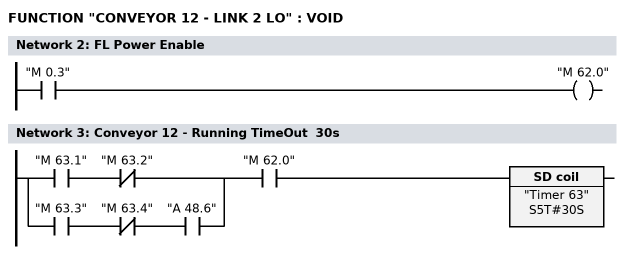

      A     "M 0.3";
      =     "M 62.0";
NETWORK
TITLE =Conveyor 12 - Running TimeOut  30s

      A(    ;
      A     "M 63.1";
      AN    "M 63.2";
      O     ;
      A     "M 63.3";
      AN    "M 63.4";
      A     "A 48.6";
      )     ;
      A     "M 62.0";
      L     S5T#30S;
      SD    "Timer 63";
NETWORK
TITLE =Conveyor 12 - Steps Register - Reset

      A(    ;
      A     "M 63.1";
      AN    "M 63.2";
      A     "Timer 63";
      O     "M 63.4";
      )     ;
      A     "M 62.0";
      JC    M001;
      JU    M002;

M001: L     W#16#0;
      T     "MW 63";
      T     "MB 65";

M002: NOP   0;
NETWORK
TITLE =Step 13N1 - Power On
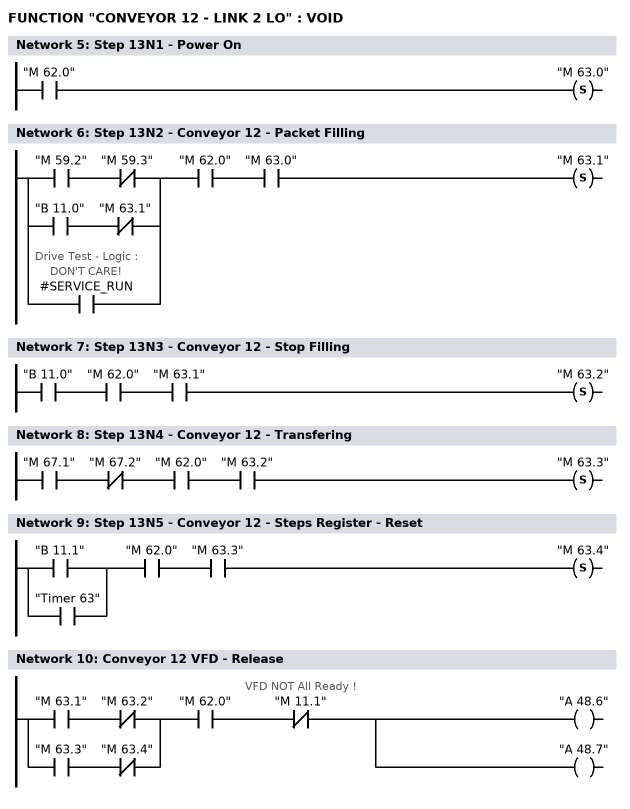

      A     "M 62.0";
      S     "M 63.0";
NETWORK
TITLE =Step 13N2 - Conveyor 12 - Packet Filling

      A(    ;
      A     "M 59.2";
      AN    "M 59.3";
      O     ;
      A     "B 11.0";
      AN    "M 63.1";
      )     ;
      O     #SERVICE_RUN; // Drive Test - Logic : DON'T CARE!
      A     "M 62.0";
      A     "M 63.0";
      S     "M 63.1";
NETWORK
TITLE =Step 13N3 - Conveyor 12 - Stop Filling

      A     "B 11.0";
      A     "M 62.0";
      A     "M 63.1";
      S     "M 63.2";
NETWORK
TITLE =Step 13N4 - Conveyor 12 - Transfering

      A     "M 67.1";
      AN    "M 67.2";
      A     "M 62.0";
      A     "M 63.2";
      S     "M 63.3";
NETWORK
TITLE =Step 13N5 - Conveyor 12 - Steps Register - Reset

      A(    ;
      O     "B 11.1";
      O     "Timer 63";
      )     ;
      A     "M 62.0";
      A     "M 63.3";
      S     "M 63.4";
NETWORK
TITLE =Conveyor 12 VFD - Release

      A(    ;
      A     "M 63.1";
      AN    "M 63.2";
      O     ;
      A     "M 63.3";
      AN    "M 63.4";
      )     ;
      A     "M 62.0";
      AN    "M 11.1"; // VFD NOT All Ready !
      =     "A 48.6";
      =     "A 48.7";
END_FUNCTION

FUNCTION "CONVEYOR 13 - DELIV. LO" : VOID
TITLE =Conveyor 13 - Delivery First Level
NAME : POS_15_L
VERSION : 0.0


VAR_TEMP
  MAIN_SERVICE_2_SW : BOOL ;
  SERVICE_RUN : BOOL ;
  BARRIER_BLINKER : BOOL ;	//Feeder Safety Light Barrier
END_VAR
BEGIN
NETWORK
TITLE =Conveyor 13 - Service

      A     "HMI_DB".ALL_SERVICE_ENABLE_SW;
      A     "HMI_DB".CONVEYOR_11_SERVICE_SW;
      A     "HMI_DB".SERVICE_SW_2_STATUS;
      =     #MAIN_SERVICE_2_SW;
//;
      A     #MAIN_SERVICE_2_SW;
      O     "M 66.1";
      JNB   CO13;
//;
      A     "HMI_DB".HMI_CONVEYOR_13_TEST_SSW;
      =     #SERVICE_RUN;
//;
      AN    #MAIN_SERVICE_2_SW;
      R     "HMI_DB".HMI_CONVEYOR_13_TEST_SSW;

CO13: R     #SERVICE_RUN;
      FP    "FP 148.2";
      =     "M 66.1";
NETWORK
TITLE =Delivery Conveyor 13 - Running TimeOut  30s
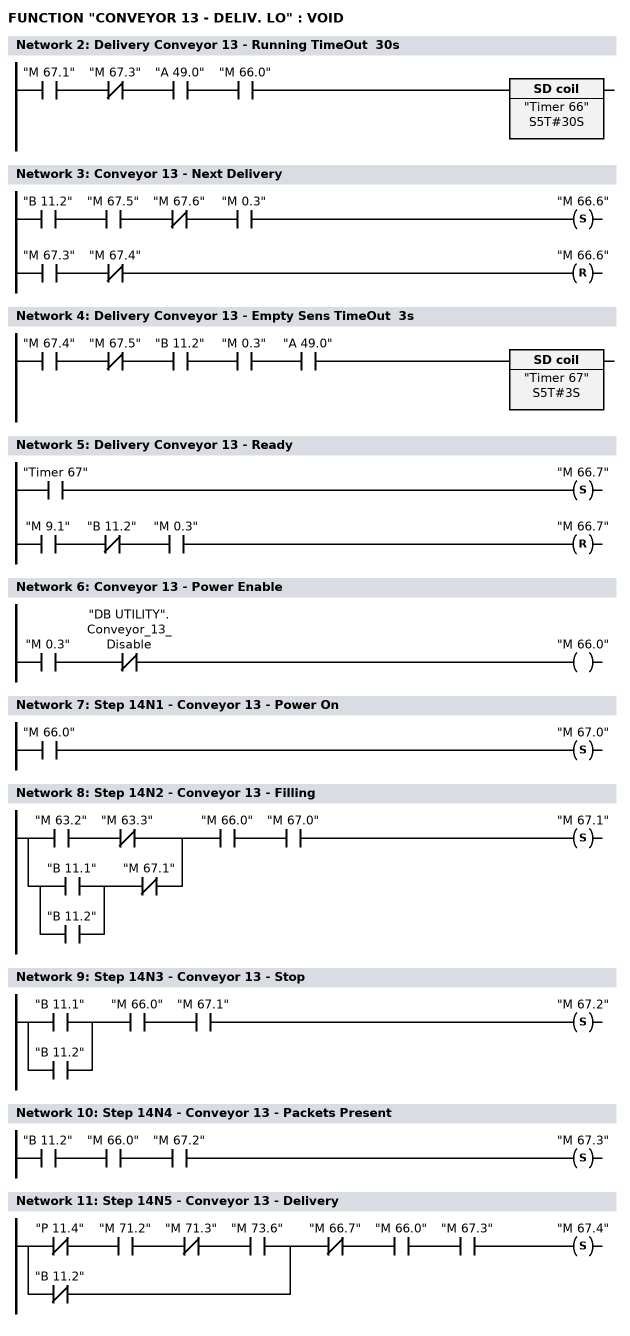

      A     "M 67.1";
      AN    "M 67.3";
      A     "A 49.0";
      A     "M 66.0";
      L     S5T#30S;
      SD    "Timer 66";
NETWORK
TITLE =Conveyor 13 - Next Delivery

      A     "B 11.2";
      A     "M 67.5";
      AN    "M 67.6";
      A     "M 0.3";
      S     "M 66.6";
//;
      A     "M 67.3";
      AN    "M 67.4";
      R     "M 66.6";
NETWORK
TITLE =Delivery Conveyor 13 - Empty Sens TimeOut  3s

      A     "M 67.4";
      AN    "M 67.5";
      A     "B 11.2";
      A     "M 0.3";
      A     "A 49.0";
      L     S5T#3S;
      SD    "Timer 67";
NETWORK
TITLE =Delivery Conveyor 13 - Ready

      A     "Timer 67";
      S     "M 66.7";
//;
      A     "M 9.1";
      AN    "B 11.2";
      A     "M 0.3";
      R     "M 66.7";
NETWORK
TITLE =Conveyor 13 - Power Enable

      A     "M 0.3";
      AN    "DB UTILITY".Conveyor_13_Disable;
      =     "M 66.0";
NETWORK
TITLE =Step 14N1 - Conveyor 13 - Power On

      A     "M 66.0";
      S     "M 67.0";
NETWORK
TITLE =Step 14N2 - Conveyor 13 - Filling

      A(    ;
      A     "M 63.2";
      AN    "M 63.3";
      O     ;
      A(    ;
      O     "B 11.1";
      O     "B 11.2";
      )     ;
//      O     #SERVICE_RUN
      AN    "M 67.1";
      )     ;
      A     "M 66.0";
      A     "M 67.0";
      S     "M 67.1";
NETWORK
TITLE =Step 14N3 - Conveyor 13 - Stop

      A(    ;
      O     "B 11.1";
      O     "B 11.2";
      )     ;
      A     "M 66.0";
      A     "M 67.1";
      S     "M 67.2";
NETWORK
TITLE =Step 14N4 - Conveyor 13 - Packets Present

      A     "B 11.2";
      A     "M 66.0";
      A     "M 67.2";
      S     "M 67.3";
NETWORK
TITLE =Step 14N5 - Conveyor 13 - Delivery

      A(    ;
      AN    "P 11.4";
      A     "M 71.2";
      AN    "M 71.3";
      A     "M 73.6";
      ON    "B 11.2";
      )     ;
      AN    "M 66.7";
      A     "M 66.0";
      A     "M 67.3";
      S     "M 67.4";
NETWORK
TITLE =Write 1 to Steps 0-3 Byte Register MB67

      A(    ;
      O     "M 66.6";
      O     "M 66.7";
      )     ;
      A     "M 67.4";
      A     "M 66.0";
      JC    M001;
      JU    M002;

M001: L     2#1111;
      T     "MB 67";

M002: NOP   0;
NETWORK
TITLE =Step 14N6 - Conveyor 13 - Delivery Done
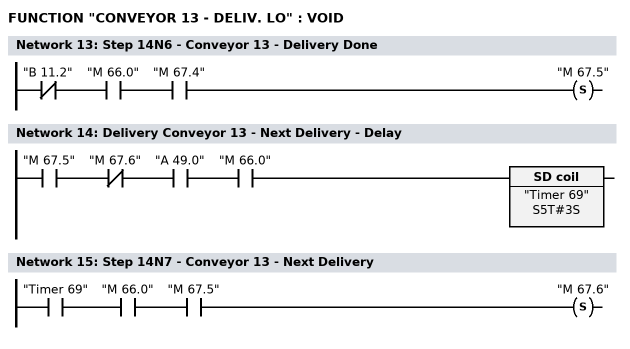

      AN    "B 11.2";
      A     "M 66.0";
      A     "M 67.4";
      S     "M 67.5";
NETWORK
TITLE =Delivery Conveyor 13 - Next Delivery - Delay

      A     "M 67.5";
      AN    "M 67.6";
      A     "A 49.0";
      A     "M 66.0";
      L     S5T#3S;
      SD    "Timer 69";
NETWORK
TITLE =Step 14N7 - Conveyor 13 - Next Delivery

      A     "Timer 69";
      A     "M 66.0";
      A     "M 67.5";
      S     "M 67.6";
NETWORK
TITLE =Steps Register - Reset

      A(    ;
      O     "M 67.6";
      O     "Timer 66";
      )     ;
      A     "M 66.0";
      JC    M003;
      JU    M004;

M003: L     2#0;
      T     "MW 67";

M004: NOP   0;
NETWORK
TITLE =Conveyor 13 VFD - Release
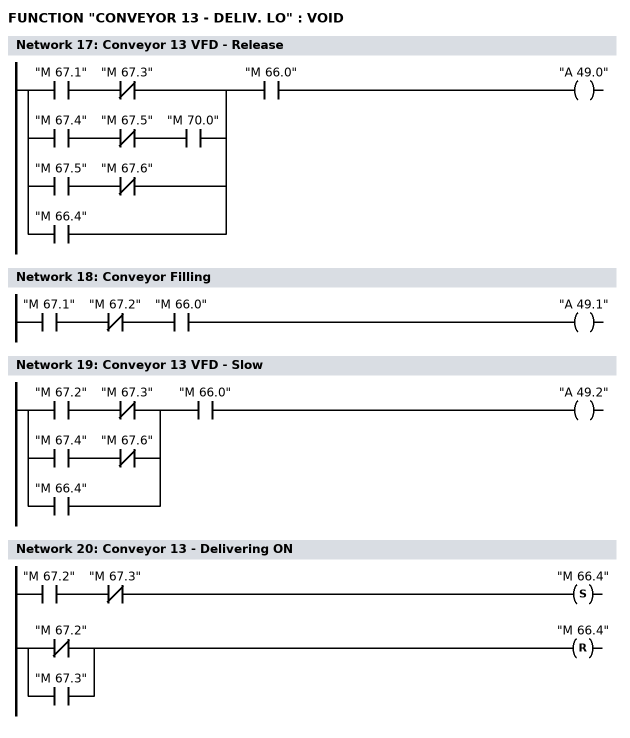

      A(    ;
      A     "M 67.1";
      AN    "M 67.3";
      O     ;
      A     "M 67.4";
      AN    "M 67.5";
      A     "M 70.0";
      O     ;
      A     "M 67.5";
      AN    "M 67.6";
      O     "M 66.4";
      )     ;
      A     "M 66.0";
      =     "A 49.0";
NETWORK
TITLE =Conveyor Filling

      A     "M 67.1";
      AN    "M 67.2";
      A     "M 66.0";
      =     "A 49.1";
NETWORK
TITLE =Conveyor 13 VFD - Slow

      A(    ;
      A     "M 67.2";
      AN    "M 67.3";
      O     ;
      A     "M 67.4";
      AN    "M 67.6";
      O     "M 66.4";
      )     ;
      A     "M 66.0";
      =     "A 49.2";
NETWORK
TITLE =Conveyor 13 - Delivering ON

      A     "M 67.2";
      AN    "M 67.3";
      S     "M 66.4";
//;
      A(    ;
      ON    "M 67.2";
      O     "M 67.3";
      )     ;
      R     "M 66.4";
END_FUNCTION

FUNCTION "LOADER FINGERS" : VOID
TITLE =Feeder Fingers
//
NAME : FEEDER
VERSION : 0.0


VAR_TEMP
  MAIN_SERVICE_3_SW : BOOL ;
  FEEDER_SERVICE_SW : BOOL ;
  FINGERS_SERVICE_SW : BOOL ;
  LIGHT_BARRIER : BOOL ;
  FINGERS_EXTEND : BOOL ;
  FINGERS_RETRACT : BOOL ;
  FINGERS_TILT : BOOL ;
  BELT_ON : BOOL ;
  INITIALISATION : BOOL ;
END_VAR
BEGIN
NETWORK
TITLE =Light Barrier Buffer
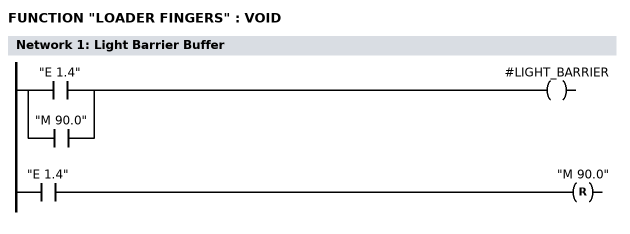

      A     "E 1.4";
      O     "M 90.0";
      =     #LIGHT_BARRIER;
//;
      A     "E 1.4";
      R     "M 90.0";
NETWORK
TITLE =Feeder Service

      A     "HMI_DB".ALL_SERVICE_ENABLE_SW;
      A     "HMI_DB".LOADER_SERVICE_ENABLE_SW;
      A     "HMI_DB".SERVICE_SW_3_STATUS;
      =     #MAIN_SERVICE_3_SW;
//;
      A     #MAIN_SERVICE_3_SW;
      O     "M 70.7";
      JNB   FEED;
      A     "HMI_DB".LOADER_LIFT_SERVICE_SSW;
      =     #FEEDER_SERVICE_SW;
//;
      A     #FEEDER_SERVICE_SW;
      A     "HMI_DB".LOADER_FING_SERVICE_SSW;
      =     #FINGERS_SERVICE_SW;
      =     "DB UTILITY".Conveyor_13_Disable;
      =     "DB UTILITY".Conveyor_23_Disable;
//;
      A     #FEEDER_SERVICE_SW;
      A     #FINGERS_SERVICE_SW;
      A     "HMI_DB".FINGER_EXTEND_TEST_PB;
      AN    #FINGERS_RETRACT;
      =     #FINGERS_EXTEND;
//;
      A     #FEEDER_SERVICE_SW;
      A     #FINGERS_SERVICE_SW;
      A     "HMI_DB".FINGER_RETRACT_TEST_PB;
      AN    #FINGERS_EXTEND;
      =     #FINGERS_RETRACT;
//;
      A     #FEEDER_SERVICE_SW;
      A     #FINGERS_SERVICE_SW;
      A     "HMI_DB".FINGER_BELT_TEST_SW;
      =     #BELT_ON;
//;
      A     #FEEDER_SERVICE_SW;
      A     #FINGERS_SERVICE_SW;
      A     "HMI_DB".FINGER_TILT_TEST_PB;
      =     #FINGERS_TILT;
//;
      AN    #MAIN_SERVICE_3_SW;
      ON    #FEEDER_SERVICE_SW;
      R     "HMI_DB".LOADER_FING_SERVICE_SSW;
      R     "HMI_DB".LOADER_LIFT_SERVICE_SSW;
      R     "HMI_DB".FINGER_RETRACT_TEST_PB;
      R     "HMI_DB".FINGER_EXTEND_TEST_PB;
      R     "HMI_DB".FINGER_TILT_TEST_PB;
      R     "HMI_DB".FINGER_BELT_TEST_SW;

FEED: R     #FEEDER_SERVICE_SW;
      R     #FINGERS_SERVICE_SW;
      R     #FINGERS_EXTEND;
      R     #FINGERS_RETRACT;
      R     #FINGERS_TILT;
      FP    "FP 159.7";
      =     "M 70.7";
//;
      A     "HMI_DB".SERVICE_INIT_PB;
      A     #FEEDER_SERVICE_SW;
      A     #MAIN_SERVICE_3_SW;
      =     #INITIALISATION;
NETWORK
TITLE =Feeder - Power Enable
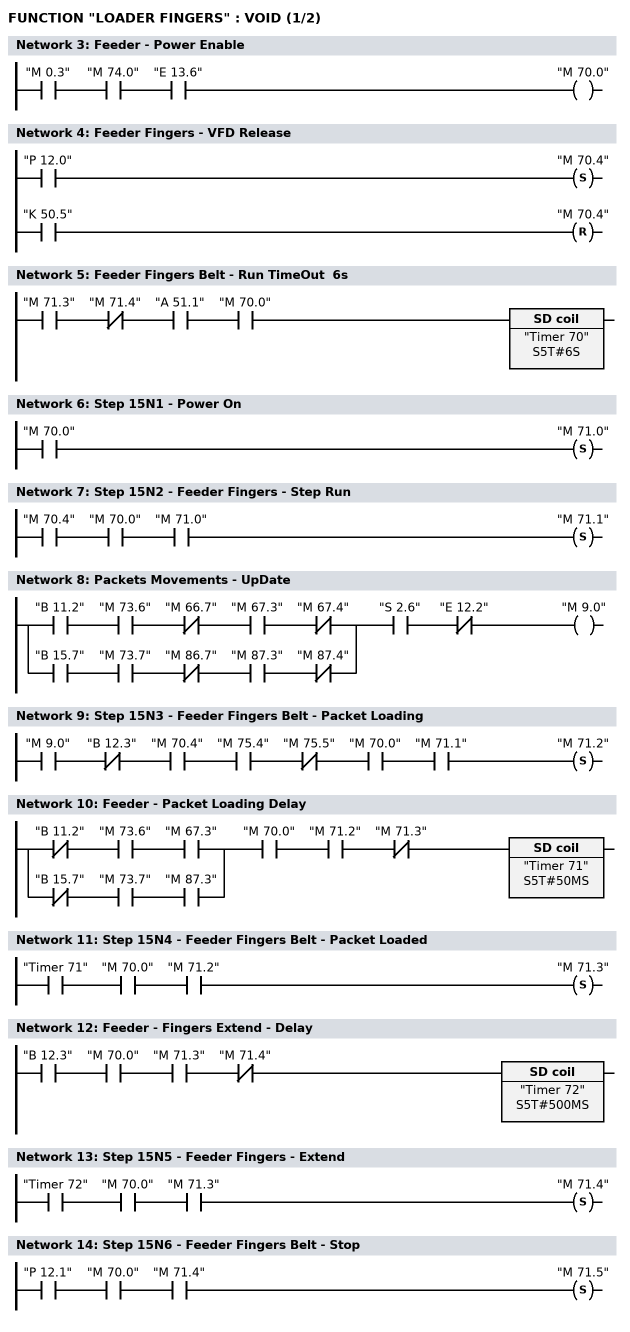

      A     "M 0.3";
      A     "M 74.0";
      A     "E 13.6";
      =     "M 70.0";
NETWORK
TITLE =Feeder Fingers - VFD Release

      A     "P 12.0";
      S     "M 70.4";
//;
      A     "K 50.5";
      R     "M 70.4";
NETWORK
TITLE =Feeder Fingers Belt - Run TimeOut  6s

      A     "M 71.3";
      AN    "M 71.4";
      A     "A 51.1";
      A     "M 70.0";
      L     S5T#6S;
      SD    "Timer 70";
NETWORK
TITLE =Step 15N1 - Power On

      A     "M 70.0";
      S     "M 71.0";
NETWORK
TITLE =Step 15N2 - Feeder Fingers - Step Run

      A     "M 70.4";
      A     "M 70.0";
      A     "M 71.0";
      S     "M 71.1";
NETWORK
TITLE =Packets Movements - UpDate

      A(    ;
      A     "B 11.2";
      A     "M 73.6";
      AN    "M 66.7";
      A     "M 67.3";
      AN    "M 67.4";
      O     ;
      A     "B 15.7";
      A     "M 73.7";
      AN    "M 86.7";
      A     "M 87.3";
      AN    "M 87.4";
      )     ;
      A     "S 2.6";
      AN    "E 12.2";
      =     "M 9.0";
NETWORK
TITLE =Step 15N3 - Feeder Fingers Belt - Packet Loading

      A     "M 9.0";
      AN    "B 12.3";
      A     "M 70.4";
      A     "M 75.4";
      AN    "M 75.5";
      A     "M 70.0";
      A     "M 71.1";
      S     "M 71.2";
NETWORK
TITLE =Feeder - Packet Loading Delay

      A(    ;
      AN    "B 11.2";
      A     "M 73.6";
      A     "M 67.3";
      O     ;
      AN    "B 15.7";
      A     "M 73.7";
      A     "M 87.3";
      )     ;
      A     "M 70.0";
      A     "M 71.2";
      AN    "M 71.3";
      L     S5T#50MS;
      SD    "Timer 71";
NETWORK
TITLE =Step 15N4 - Feeder Fingers Belt - Packet Loaded

      A     "Timer 71";
      A     "M 70.0";
      A     "M 71.2";
      S     "M 71.3";
NETWORK
TITLE =Feeder - Fingers Extend - Delay

      A     "B 12.3";
      A     "M 70.0";
      A     "M 71.3";
      AN    "M 71.4";
      L     S5T#500MS;
      SD    "Timer 72";
NETWORK
TITLE =Step 15N5 - Feeder Fingers - Extend

      A     "Timer 72";
      A     "M 70.0";
      A     "M 71.3";
      S     "M 71.4";
NETWORK
TITLE =Step 15N6 - Feeder Fingers Belt - Stop

      A     "P 12.1";
      A     "M 70.0";
      A     "M 71.4";
      S     "M 71.5";
NETWORK
TITLE =Step 15N7 - Feeder Fingers Tilt - Ready
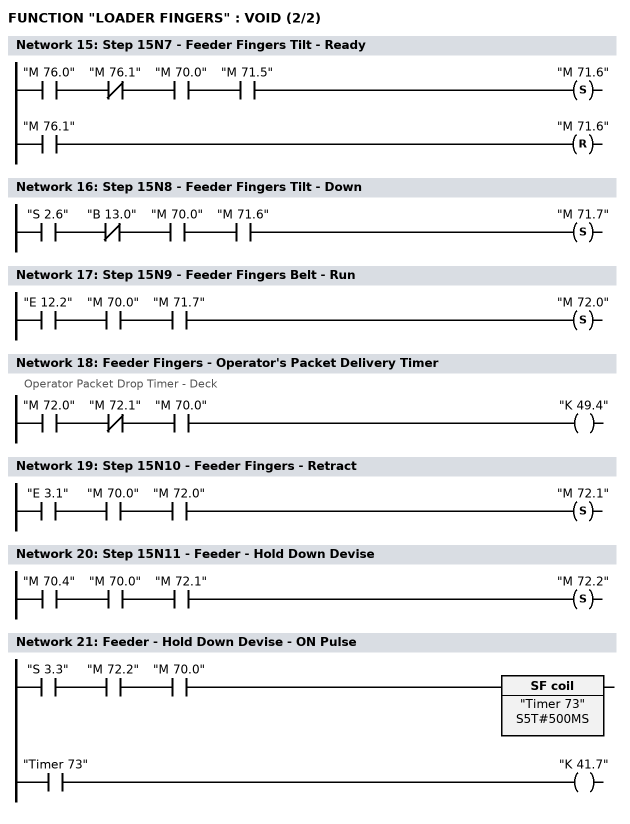

      A     "M 76.0";
      AN    "M 76.1";
      A     "M 70.0";
      A     "M 71.5";
      S     "M 71.6";
//;
      O     "M 76.1";
      R     "M 71.6";
NETWORK
TITLE =Step 15N8 - Feeder Fingers Tilt - Down

      A     "S 2.6";
      AN    "B 13.0";
      A     "M 70.0";
      A     "M 71.6";
      S     "M 71.7";
NETWORK
TITLE =Step 15N9 - Feeder Fingers Belt - Run

      A     "E 12.2";
      A     "M 70.0";
      A     "M 71.7";
      S     "M 72.0";
NETWORK
TITLE =Feeder Fingers - Operator's Packet Delivery Timer
//Operator Packet Drop Timer - Deck
      A     "M 72.0";
      AN    "M 72.1";
      A     "M 70.0";
      =     "K 49.4";
NETWORK
TITLE =Step 15N10 - Feeder Fingers - Retract

      A     "E 3.1";
      A     "M 70.0";
      A     "M 72.0";
      S     "M 72.1";
NETWORK
TITLE =Step 15N11 - Feeder - Hold Down Devise

      A     "M 70.4";
      A     "M 70.0";
      A     "M 72.1";
      S     "M 72.2";
NETWORK
TITLE =Feeder - Hold Down Devise - ON Pulse

      A     "S 3.3";
      A     "M 72.2";
      A     "M 70.0";
      L     S5T#500MS;
      SF    "Timer 73";

      A     "Timer 73";
      =     "K 41.7";
NETWORK
TITLE =Feeder Fingers - Steps Chain Register Reset

      A(    ;
      ON    "M 75.0";
      O     "M 72.2";
      O     "Timer 70";
      O     #FEEDER_SERVICE_SW;
      )     ;
      JC    M001;
      JU    M002;

M001: L     2#0;
      T     "MW 71";

M002: NOP   0;
NETWORK
TITLE =Feeder Fingers - Fingers Retract
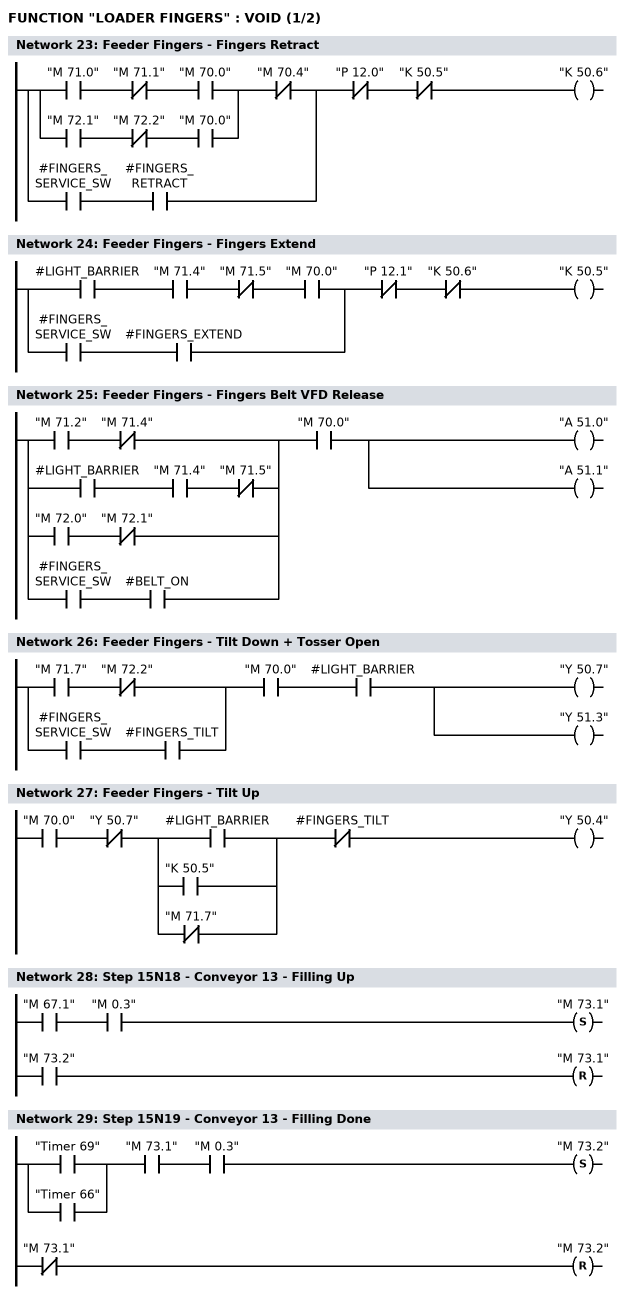

      A(    ;
      A(    ;
      A     "M 71.0";
      AN    "M 71.1";
      A     "M 70.0";
      O     ;
      A     "M 72.1";
      AN    "M 72.2";
      A     "M 70.0";
      )     ;
      AN    "M 70.4";
      O     ;
      A     #FINGERS_SERVICE_SW;
      A     #FINGERS_RETRACT;
      )     ;
      AN    "P 12.0";
      AN    "K 50.5";
      =     "K 50.6";
NETWORK
TITLE =Feeder Fingers - Fingers Extend

      A(    ;
      A     #LIGHT_BARRIER;
      A     "M 71.4";
      AN    "M 71.5";
      A     "M 70.0";
      O     ;
      A     #FINGERS_SERVICE_SW;
      A     #FINGERS_EXTEND;
      )     ;
      AN    "P 12.1";
      AN    "K 50.6";
      =     "K 50.5";
NETWORK
TITLE =Feeder Fingers - Fingers Belt VFD Release

      A(    ;
      A     "M 71.2";
      AN    "M 71.4";
      O     ;
      A     #LIGHT_BARRIER;
      A     "M 71.4";
      AN    "M 71.5";
      O     ;
      A     "M 72.0";
      AN    "M 72.1";
      O     ;
      A     #FINGERS_SERVICE_SW;
      A     #BELT_ON;
      )     ;
      A     "M 70.0";
      =     "A 51.0";
      =     "A 51.1";
NETWORK
TITLE =Feeder Fingers - Tilt Down + Tosser Open

      A(    ;
      A     "M 71.7";
      AN    "M 72.2";
      O     ;
      A     #FINGERS_SERVICE_SW;
      A     #FINGERS_TILT;
      )     ;
      A     "M 70.0";
      A     #LIGHT_BARRIER;
      =     "Y 50.7";
      =     "Y 51.3";
NETWORK
TITLE =Feeder Fingers - Tilt Up

      A     "M 70.0";
      AN    "Y 50.7";
      A(    ;
      O     #LIGHT_BARRIER;
      O     "K 50.5";
      ON    "M 71.7";
      AN    #FINGERS_TILT;
      )     ;
      =     "Y 50.4";
NETWORK
TITLE =Step 15N18 - Conveyor 13 - Filling Up

      A     "M 67.1";
      A     "M 0.3";
      S     "M 73.1";
//;
      A     "M 73.2";
      R     "M 73.1";
NETWORK
TITLE =Step 15N19 - Conveyor 13 - Filling Done

      A(    ;
      O     "Timer 69";
      O     "Timer 66";
      )     ;
      A     "M 73.1";
      A     "M 0.3";
      S     "M 73.2";
//;
      AN    "M 73.1";
      R     "M 73.2";
NETWORK
TITLE =Step 15N20 - Conveyor 23 - Filling Up
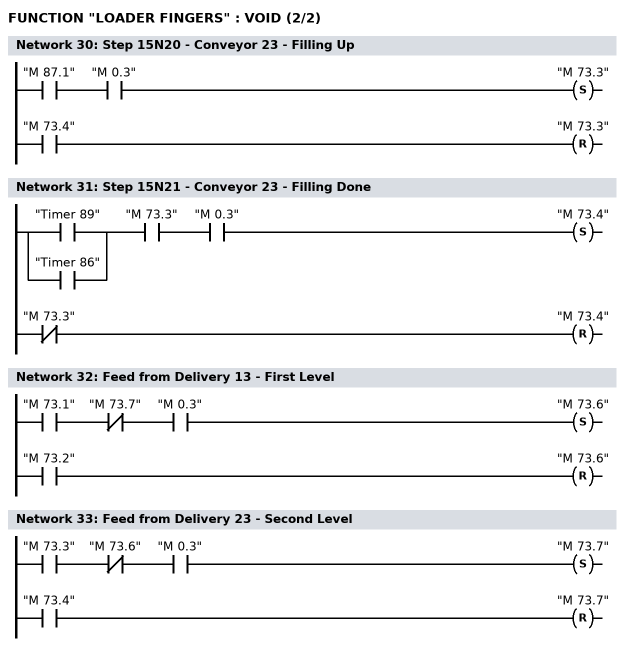

      A     "M 87.1";
      A     "M 0.3";
      S     "M 73.3";
//;
      A     "M 73.4";
      R     "M 73.3";
NETWORK
TITLE =Step 15N21 - Conveyor 23 - Filling Done

      A(    ;
      O     "Timer 89";
      O     "Timer 86";
      )     ;
      A     "M 73.3";
      A     "M 0.3";
      S     "M 73.4";
//;
      AN    "M 73.3";
      R     "M 73.4";
NETWORK
TITLE =Feed from Delivery 13 - First Level

      A     "M 73.1";
      AN    "M 73.7";
      A     "M 0.3";
      S     "M 73.6";
//;
      A     "M 73.2";
      R     "M 73.6";
NETWORK
TITLE =Feed from Delivery 23 - Second Level

      A     "M 73.3";
      AN    "M 73.6";
      A     "M 0.3";
      S     "M 73.7";
//;
      A     "M 73.4";
      R     "M 73.7";
END_FUNCTION

FUNCTION "LOADER LIFT" : VOID
TITLE =Feeder Lift   Pos. 16
//
NAME : FEEDER
VERSION : 0.0


VAR_TEMP
  MAIN_SERVICE_3_SW : BOOL ;
  FEEDER_SW : BOOL ;
  FEEDER_SERVICE_SW : BOOL ;
  LIGHT_BARRIER : BOOL ;
  FEEDER_LIFT_TOP_PB : BOOL ;
  FEEDER_LIFT_UP_PB : BOOL ;
  FEEDER_LIFT_DN_PB : BOOL ;
  FEEDER_LIFT_JOG_UP : BOOL ;
  FEEDER_LIFT_JOG_DN : BOOL ;
END_VAR
BEGIN
NETWORK
TITLE =Light Barrier Buffer
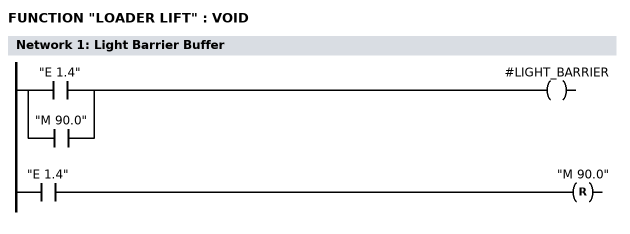

      A     "E 1.4";
      O     "M 90.0";
      =     #LIGHT_BARRIER;
//;
      A     "E 1.4";
      R     "M 90.0";
NETWORK
TITLE =Feeder Service

      A     "HMI_DB".ALL_SERVICE_ENABLE_SW;
      A     "HMI_DB".LOADER_SERVICE_ENABLE_SW;
      A     "HMI_DB".SERVICE_SW_3_STATUS;
      =     #MAIN_SERVICE_3_SW;
//;
      A     #MAIN_SERVICE_3_SW;
      O     "M 74.7";
      JNB   FEED;
      A     "HMI_DB".LOADER_LIFT_SERVICE_SSW;
      =     #FEEDER_SERVICE_SW;
      S     "DB UTILITY".Conveyor_13_Disable;
      S     "DB UTILITY".Conveyor_23_Disable;
      R     "M 74.2";
//;
      A     #FEEDER_SERVICE_SW;
      A     "HMI_DB".LOADER_LIFT_TOP_PB;
      =     #FEEDER_LIFT_TOP_PB;
//;
      A     #FEEDER_SERVICE_SW;
      A     "HMI_DB".LOADER_LIFT_UP_PB;
      =     #FEEDER_LIFT_UP_PB;
//;
      A     #FEEDER_SERVICE_SW;
      A     "HMI_DB".LOADER_LIFT_DN_PB;
      =     #FEEDER_LIFT_DN_PB;
//;
      AN    #MAIN_SERVICE_3_SW;
      ON    #FEEDER_SERVICE_SW;
      R     "HMI_DB".LOADER_FING_SERVICE_SSW;
      R     "HMI_DB".LOADER_LIFT_SERVICE_SSW;
      R     "HMI_DB".LOADER_LIFT_TOP_PB;
      R     "HMI_DB".LOADER_LIFT_UP_PB;
      R     "HMI_DB".LOADER_LIFT_DN_PB;
      R     "DB UTILITY".Conveyor_13_Disable;
      R     "DB UTILITY".Conveyor_23_Disable;

FEED: R     #FEEDER_SERVICE_SW;
      R     #FEEDER_LIFT_TOP_PB;
      R     #FEEDER_LIFT_UP_PB;
      R     #FEEDER_LIFT_DN_PB;
      FP    "FP 159.6";
      =     "M 74.7";
NETWORK
TITLE =Automatic Trigger
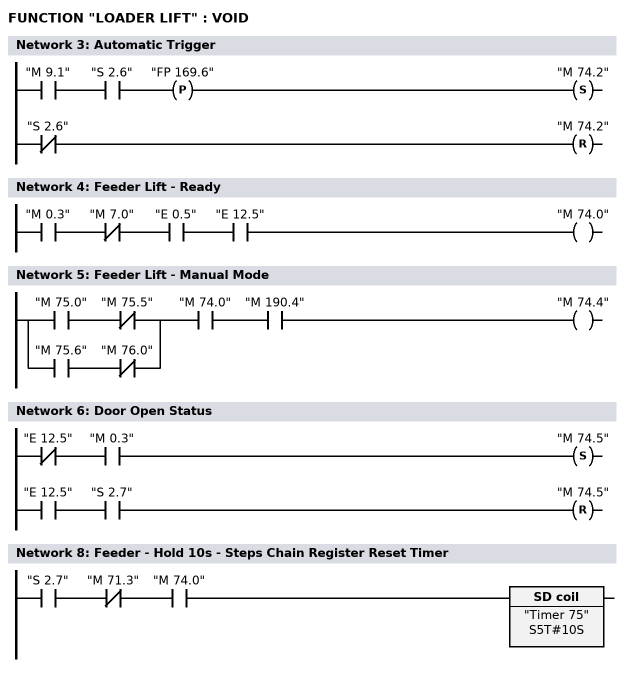

      O     "M 9.1";
      A     "S 2.6";
      FP    "FP 169.6";
      S     "M 74.2";
//;
      AN    "S 2.6";
      R     "M 74.2";
NETWORK
TITLE =Feeder Lift - Ready

      A     "M 0.3";
      AN    "M 7.0";
      A     "E 0.5";
      A     "E 12.5";
      =     "M 74.0";
NETWORK
TITLE =Feeder Lift - Manual Mode

      A(    ;
      A     "M 75.0";
      AN    "M 75.5";
      O     ;
      A     "M 75.6";
      AN    "M 76.0";
      )     ;
      A     "M 74.0";
      A     "M 190.4";
      =     "M 74.4";
NETWORK
TITLE =Door Open Status

      AN    "E 12.5";
      A     "M 0.3";
      S     "M 74.5";
//;
      A     "E 12.5";
      A     "S 2.7";
      R     "M 74.5";
NETWORK
TITLE =Fault Reset Status        X121     transfered to FC 212 Net 79
//      A(
//      O     "M 54.7"
//      O     "M 66.7"
//      O     "M 86.7"
//      )
//      A     "M 145.0"
//      O     "M 74.5"
//      O     "Timer 0"
//      =     "H 40.3"
//
//is transfered to FC 212 Net 79


NETWORK
TITLE =Feeder - Hold 10s - Steps Chain Register Reset Timer

      A     "S 2.7";
      AN    "M 71.3";
      A     "M 74.0";
      L     S5T#10S;
      SD    "Timer 75";
NETWORK
TITLE =Feeder - All Register Reset

      A(    ;
      A     "M 190.4";
      A     "M 171.4";
      A     "M 171.5";
      O     "Timer 75";
      )     ;
      A     "M 74.0";
      JC    M001;
      JU    M002;

M001: L     2#0;
      T     "MW 71";
      T     "MW 75";

M002: NOP   0;
NETWORK
TITLE =Step 16N1 - Power On
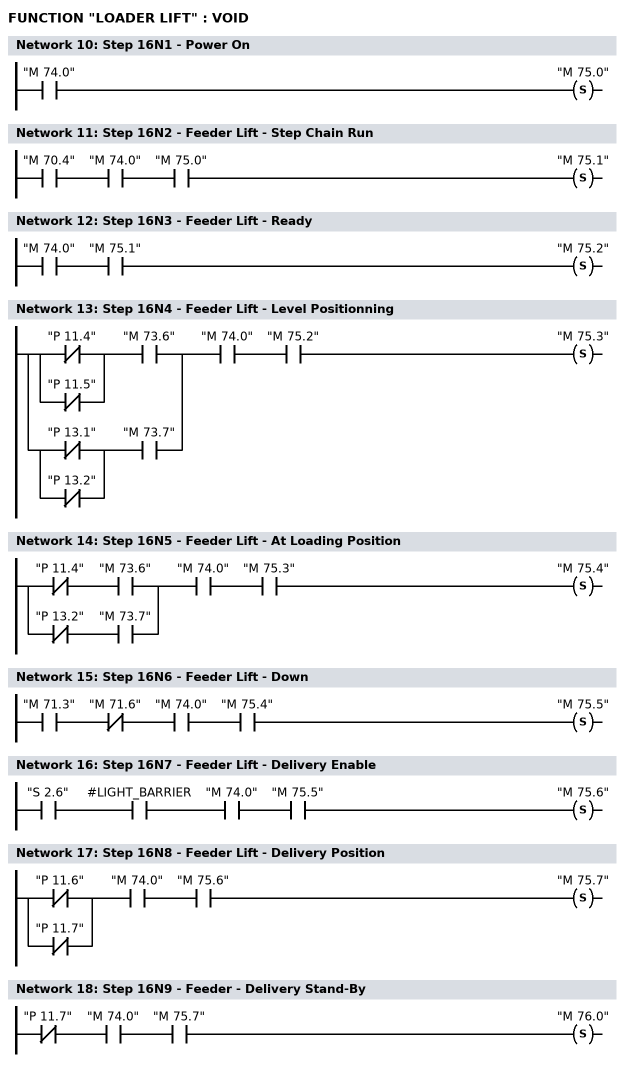

      A     "M 74.0";
      S     "M 75.0";
NETWORK
TITLE =Step 16N2 - Feeder Lift - Step Chain Run

      A     "M 70.4";
      A     "M 74.0";
      A     "M 75.0";
      S     "M 75.1";
NETWORK
TITLE =Step 16N3 - Feeder Lift - Ready

      A     "M 74.0";
      A     "M 75.1";
      S     "M 75.2";
NETWORK
TITLE =Step 16N4 - Feeder Lift - Level Positionning

      A(    ;
      A(    ;
      ON    "P 11.4";
      ON    "P 11.5";
      )     ;
      A     "M 73.6";
      O     ;
      A(    ;
      ON    "P 13.1";
      ON    "P 13.2";
      )     ;
      A     "M 73.7";
      )     ;
      A     "M 74.0";
      A     "M 75.2";
      S     "M 75.3";
NETWORK
TITLE =Step 16N5 - Feeder Lift - At Loading Position

      A(    ;
      AN    "P 11.4";
      A     "M 73.6";
      O     ;
      AN    "P 13.2";
      A     "M 73.7";
      )     ;
      A     "M 74.0";
      A     "M 75.3";
      S     "M 75.4";
NETWORK
TITLE =Step 16N6 - Feeder Lift - Down

      A     "M 71.3";
      AN    "M 71.6";
      A     "M 74.0";
      A     "M 75.4";
      S     "M 75.5";
NETWORK
TITLE =Step 16N7 - Feeder Lift - Delivery Enable

      A     "S 2.6";
      A     #LIGHT_BARRIER;
      A     "M 74.0";
      A     "M 75.5";
      S     "M 75.6";
NETWORK
TITLE =Step 16N8 - Feeder Lift - Delivery Position

      A(    ;
      ON    "P 11.6";
      ON    "P 11.7";
      )     ;
      A     "M 74.0";
      A     "M 75.6";
      S     "M 75.7";
NETWORK
TITLE =Step 16N9 - Feeder - Delivery Stand-By

      AN    "P 11.7";
      A     "M 74.0";
      A     "M 75.7";
      S     "M 76.0";
NETWORK
TITLE =Feeder Lift Steps Chain Reset by Feeder Fingers (MW71)

      A     "M 76.0";
      AN    "M 76.1";
      A(    ;
      ON    "M 71.2";
      O     "M 72.2";
      )     ;
      A     "M 74.0";
      JC    M003;
      JU    M004;

M003: L     2#0;
      T     "MW 75";

M004: NOP   0;
NETWORK
TITLE =Step 16N10 - Feeder Hold Operation (Stop) 1
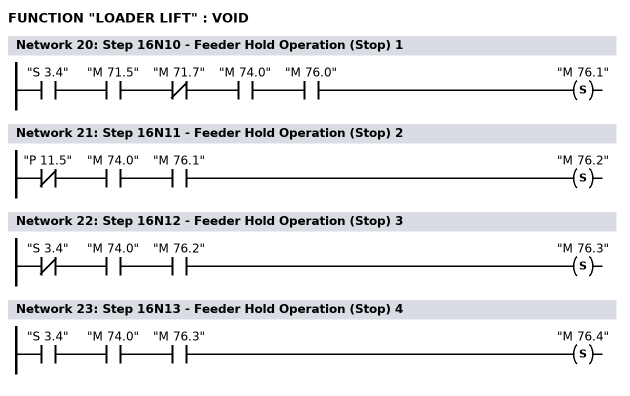

      A     "S 3.4";
      A     "M 71.5";
      AN    "M 71.7";
      A     "M 74.0";
      A     "M 76.0";
      S     "M 76.1";
NETWORK
TITLE =Step 16N11 - Feeder Hold Operation (Stop) 2

      AN    "P 11.5";
      A     "M 74.0";
      A     "M 76.1";
      S     "M 76.2";
NETWORK
TITLE =Step 16N12 - Feeder Hold Operation (Stop) 3

      AN    "S 3.4";
      A     "M 74.0";
      A     "M 76.2";
      S     "M 76.3";
NETWORK
TITLE =Step 16N13 - Feeder Hold Operation (Stop) 4

      A     "S 3.4";
      A     "M 74.0";
      A     "M 76.3";
      S     "M 76.4";
NETWORK
TITLE =Step 16N14 - Feeder Hold Operation (Stop) 4 - Fill MB76

      A     "M 76.4";
      A     "M 74.0";
      JC    M005;
      JU    M006;

M005: L     2#11111100000000;
      T     "MW 75";

M006: NOP   0;
NETWORK
TITLE =Packets Movements - UpDate
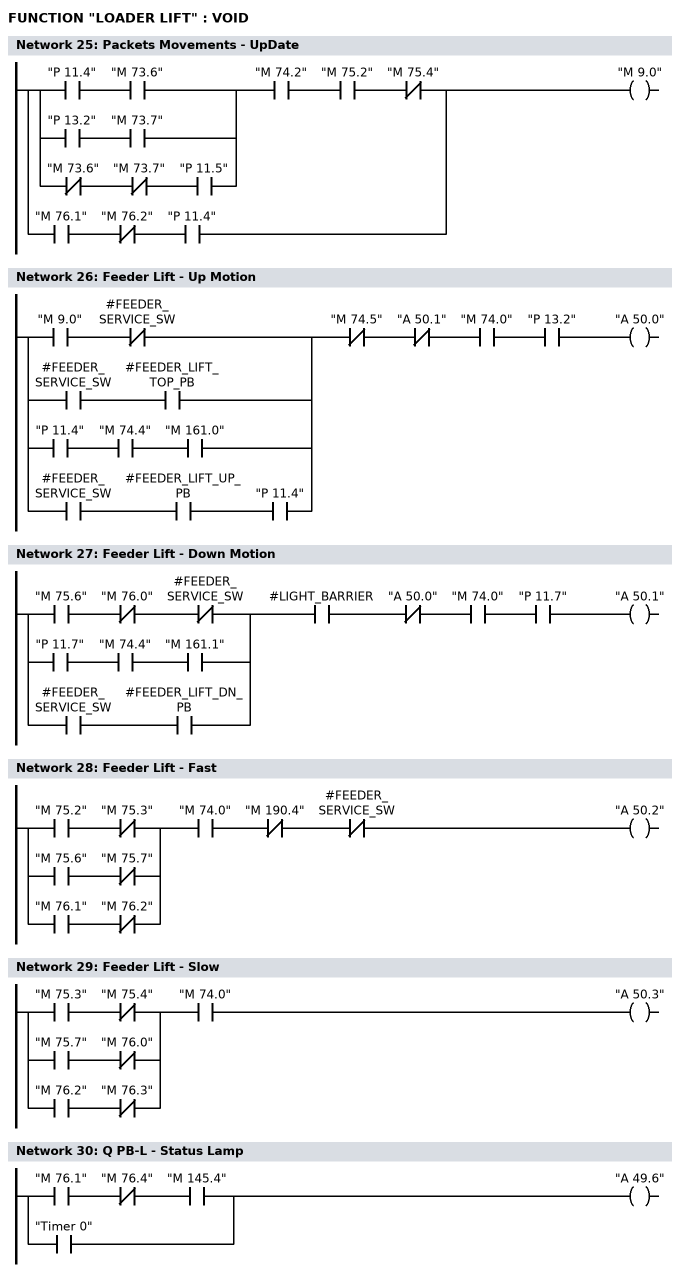

      A(    ;
      A     "P 11.4";
      A     "M 73.6";
      O     ;
      A     "P 13.2";
      A     "M 73.7";
      O     ;
      AN    "M 73.6";
      AN    "M 73.7";
      A     "P 11.5";
      )     ;
      A     "M 74.2";
      A     "M 75.2";
      AN    "M 75.4";
      O     ;
      A     "M 76.1";
      AN    "M 76.2";
      A     "P 11.4";
      =     "M 9.0";
NETWORK
TITLE =Feeder Lift - Up Motion

      A(    ;
      A     "M 9.0";
      AN    #FEEDER_SERVICE_SW;
      O     ;
      A     #FEEDER_SERVICE_SW;
      A     #FEEDER_LIFT_TOP_PB;

      O     ;
      A     "P 11.4";
      A     "M 74.4";
      A     "M 161.0";

      O     ;
      A     #FEEDER_SERVICE_SW;
      A     #FEEDER_LIFT_UP_PB;
      A     "P 11.4";
      )     ;
      AN    "M 74.5";
      AN    "A 50.1";
      A     "M 74.0";
      A     "P 13.2";
      =     "A 50.0";
NETWORK
TITLE =Feeder Lift - Down Motion

      A(    ;
      A     "M 75.6";
      AN    "M 76.0";
      AN    #FEEDER_SERVICE_SW;

      O     ;
      A     "P 11.7";
      A     "M 74.4";
      A     "M 161.1";

      O     ;
      A     #FEEDER_SERVICE_SW;
      A     #FEEDER_LIFT_DN_PB;
      )     ;
      A     #LIGHT_BARRIER;
      AN    "A 50.0";
      A     "M 74.0";
      A     "P 11.7";
      =     "A 50.1";
NETWORK
TITLE =Feeder Lift - Fast

      A(    ;
      A     "M 75.2";
      AN    "M 75.3";
      O     ;
      A     "M 75.6";
      AN    "M 75.7";
      O     ;
      A     "M 76.1";
      AN    "M 76.2";
      )     ;
      A     "M 74.0";
      AN    "M 190.4";
      AN    #FEEDER_SERVICE_SW;
      =     "A 50.2";
NETWORK
TITLE =Feeder Lift - Slow

      A(    ;
      A     "M 75.3";
      AN    "M 75.4";
      O     ;
      A     "M 75.7";
      AN    "M 76.0";
      O     ;
      A     "M 76.2";
      AN    "M 76.3";
      )     ;
      A     "M 74.0";
      =     "A 50.3";
NETWORK
TITLE =Q PB-L - Status Lamp

      A     "M 76.1";
      AN    "M 76.4";
      A     "M 145.4";
      O     "Timer 0";
      =     "A 49.6";
END_FUNCTION

FUNCTION "CONVEYOR 21 - LINK 1 HI" : VOID
TITLE =Conveyor 21 - Link 1H  Pos. 13 High Level
//
NAME : POS_13_H
VERSION : 0.0


VAR_TEMP
  MAIN_SERVICE_2_SW : BOOL ;
  SERVICE_RUN : BOOL ;
  INITIALISATION : BOOL ;
  BARRIER_BLINKER : BOOL ;
END_VAR
BEGIN
NETWORK
TITLE =Conveyor 21 - Service

      A     "HMI_DB".ALL_SERVICE_ENABLE_SW;
      A     "HMI_DB".CONVEYOR_21_SERVICE_SW;
      A     "HMI_DB".SERVICE_SW_2_STATUS;
      =     #MAIN_SERVICE_2_SW;
//;
      A     #MAIN_SERVICE_2_SW;
      O     "M 78.7";
      JNB   CO21;
//;
      A     "HMI_DB".HMI_CONVEYOR_21_TEST_SSW;
      AN    "A 48.0";
      =     #SERVICE_RUN;
      S     "DB UTILITY".Conveyor_10_Disable;
      S     "DB UTILITY".Pivot_Disable;
//;
      A     "HMI_DB".SERVICE_INIT_PB;
      =     #INITIALISATION;
//;
      AN    #MAIN_SERVICE_2_SW;
      R     "HMI_DB".HMI_CONVEYOR_21_TEST_SSW;
      R     "DB UTILITY".Conveyor_10_Disable;
      R     "DB UTILITY".Pivot_Disable;

CO21: R     #SERVICE_RUN;
      FP    "FP 148.3";
      =     "M 78.7";
NETWORK
TITLE =Power Enable
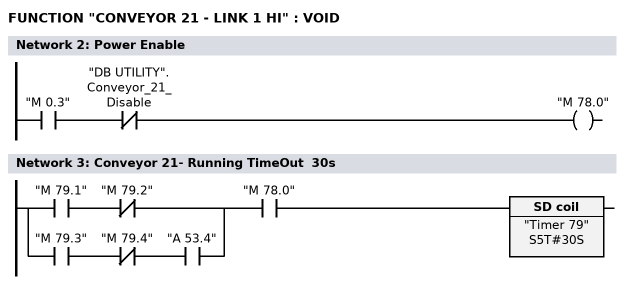

      A     "M 0.3";
      AN    "DB UTILITY".Conveyor_21_Disable;
      =     "M 78.0";
NETWORK
TITLE =Conveyor 21- Running TimeOut  30s

      A(    ;
      A     "M 79.1";
      AN    "M 79.2";
      O     ;
      A     "M 79.3";
      AN    "M 79.4";
      A     "A 53.4";
      )     ;
      A     "M 78.0";
      L     S5T#30S;
      SD    "Timer 79"; // C21 TimeOut
NETWORK
TITLE =Steps Register - Reset

      A(    ;
      A     "M 79.1"; // Filling Step
      AN    "M 79.2"; // Filling Step - Done
      A     "Timer 79"; // C21 TimeOut
      O     "M 79.4";
      O     #INITIALISATION;
      O     "DB UTILITY".Conveyor_21_Disable;
      )     ;
      A     "M 78.0";
      JC    M001;
      JU    M002;

M001: L     W#16#0;
      T     "MW 79"; // Step Register - Reset
      T     "MB 81"; // Step Register - Reset

M002: NOP   0;
NETWORK
TITLE =Step 22N1 - Power ON
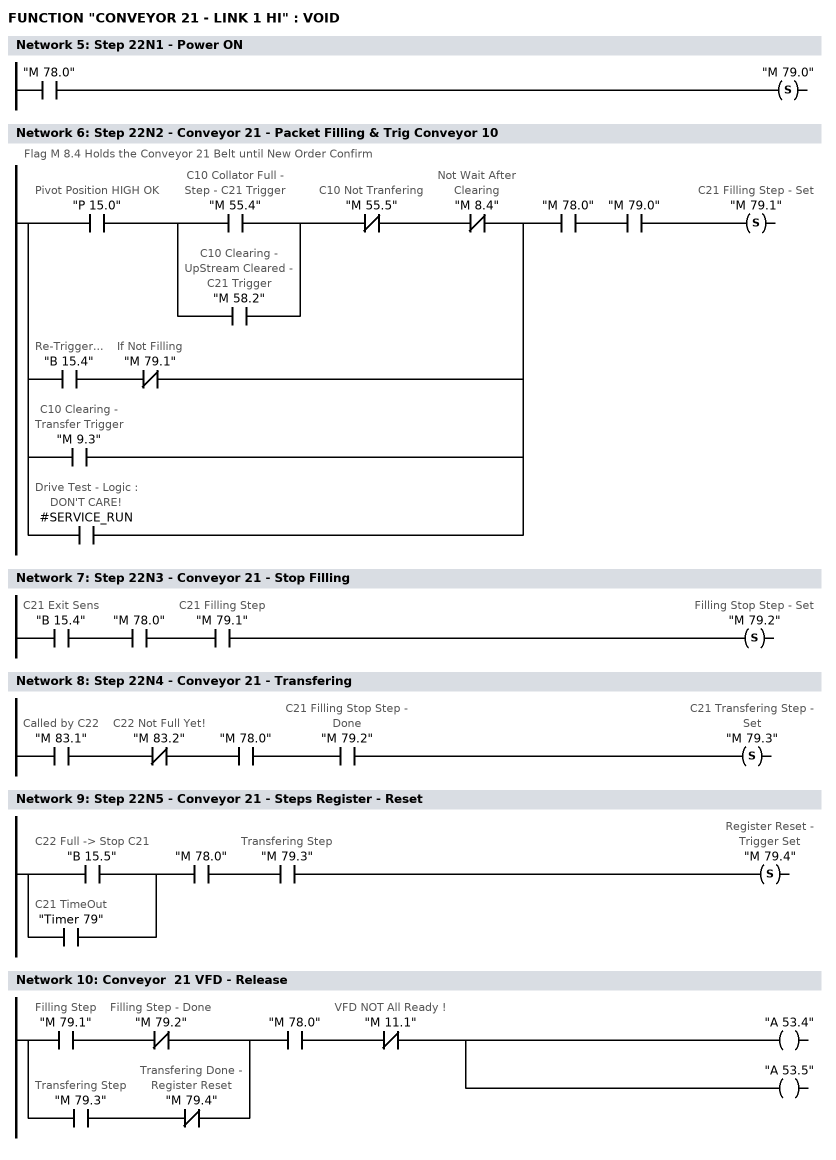

      A     "M 78.0";
      S     "M 79.0";
NETWORK
TITLE =Step 22N2 - Conveyor 21 - Packet Filling & Trig Conveyor 10
//Flag M 8.4 Holds the Conveyor 21 Belt until New Order Confirm
      A(    ;
      A     "P 15.0"; // Pivot Position HIGH OK
      A(    ;
      O     "M 55.4"; // C10 Collator Full - Step - C21 Trigger
      O     "M 58.2"; // C10 Clearing - UpStream Cleared - C21 Trigger
      )     ;
      AN    "M 55.5"; // C10 Not Tranfering
      AN    "M 8.4"; // Not Wait After Clearing
      O     ;
      A     "B 15.4"; // Re-Trigger...
      AN    "M 79.1"; // If Not Filling
      O     ;
      A     "M 9.3"; // C10 Clearing - Transfer Trigger
      )     ;
      O     #SERVICE_RUN; // Drive Test - Logic : DON'T CARE!
      A     "M 78.0";
      A     "M 79.0";
      S     "M 79.1"; // C21 Filling Step - Set
NETWORK
TITLE =Step 22N3 - Conveyor 21 - Stop Filling

      A     "B 15.4"; // C21 Exit Sens
      A     "M 78.0";
      A     "M 79.1"; // C21 Filling Step
      S     "M 79.2"; // Filling Stop Step - Set
NETWORK
TITLE =Step 22N4 - Conveyor 21 - Transfering

      A     "M 83.1"; // Called by C22
      AN    "M 83.2"; // C22 Not Full Yet!
      A     "M 78.0";
      A     "M 79.2"; // C21 Filling Stop Step - Done
      S     "M 79.3"; // C21 Transfering Step - Set
NETWORK
TITLE =Step 22N5 - Conveyor 21 - Steps Register - Reset

      A(    ;
      O     "B 15.5"; // C22 Full -> Stop C21
      O     "Timer 79"; // C21 TimeOut
      )     ;
      A     "M 78.0";
      A     "M 79.3"; // Transfering Step
      S     "M 79.4"; // Register Reset - Trigger Set
NETWORK
TITLE =Conveyor  21 VFD - Release

      A(    ;
      A     "M 79.1"; // Filling Step
      AN    "M 79.2"; // Filling Step - Done
      O     ;
      A     "M 79.3"; // Transfering Step
      AN    "M 79.4"; // Transfering Done - Register Reset
      )     ;
      A     "M 78.0";
      AN    "M 11.1"; // VFD NOT All Ready !
      =     "A 53.4";
      =     "A 53.5";
END_FUNCTION

FUNCTION "CONVEYOR 22 - LINK 2 HI" : VOID
TITLE =Conveyor 22 - Link 2H  Pos. 14 High Level
//
NAME : POS_14_H
VERSION : 0.0


VAR_TEMP
  MAIN_SERVICE_2_SW : BOOL ;
  SERVICE_RUN : BOOL ;
END_VAR
BEGIN
NETWORK
TITLE =Conveyor 22 - Service

      A     "HMI_DB".ALL_SERVICE_ENABLE_SW;
      A     "HMI_DB".CONVEYOR_21_SERVICE_SW;
      A     "HMI_DB".SERVICE_SW_2_STATUS;
      =     #MAIN_SERVICE_2_SW;
//;
      A     #MAIN_SERVICE_2_SW;
      O     "M 82.7";
      JNB   CO22;
//;
      A     "HMI_DB".HMI_CONVEYOR_22_TEST_SSW;
      =     #SERVICE_RUN;
//;
      AN    #MAIN_SERVICE_2_SW;
      R     "HMI_DB".HMI_CONVEYOR_22_TEST_SSW;

CO22: R     #SERVICE_RUN;
      FP    "FP 148.4";
      =     "M 82.7";
NETWORK
TITLE =Power Enable
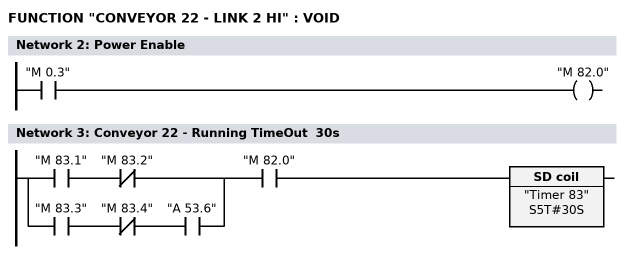

      A     "M 0.3";
      =     "M 82.0";
NETWORK
TITLE =Conveyor 22 - Running TimeOut  30s

      A(    ;
      A     "M 83.1";
      AN    "M 83.2";
      O     ;
      A     "M 83.3";
      AN    "M 83.4";
      A     "A 53.6";
      )     ;
      A     "M 82.0";
      L     S5T#30S;
      SD    "Timer 83";
NETWORK
TITLE =Conveyor 22 - Steps Register - Reset

      A(    ;
      A     "M 83.1";
      AN    "M 83.2";
      A     "Timer 83";
      O     "M 83.4";
      )     ;
      A     "M 82.0";
      JC    M001;
      JU    M002;

M001: L     W#16#0;
      T     "MW 83";
      T     "MB 85";

M002: NOP   0;
NETWORK
TITLE =Step 23N1 - Power On
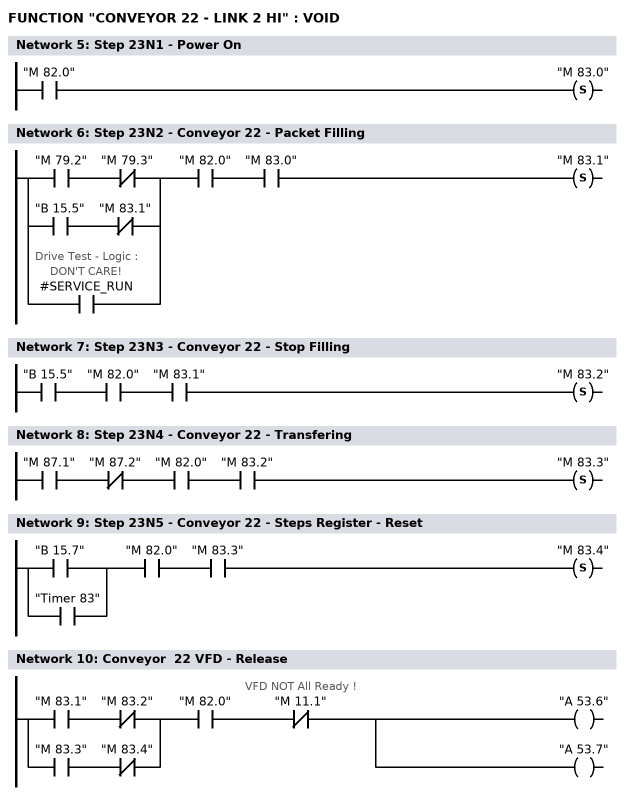

      A     "M 82.0";
      S     "M 83.0";
NETWORK
TITLE =Step 23N2 - Conveyor 22 - Packet Filling

      A(    ;
      A     "M 79.2";
      AN    "M 79.3";
      O     ;
      A     "B 15.5";
      AN    "M 83.1";
      )     ;
      O     #SERVICE_RUN; // Drive Test - Logic : DON'T CARE!
      A     "M 82.0";
      A     "M 83.0";
      S     "M 83.1";
NETWORK
TITLE =Step 23N3 - Conveyor 22 - Stop Filling

      A     "B 15.5";
      A     "M 82.0";
      A     "M 83.1";
      S     "M 83.2";
NETWORK
TITLE =Step 23N4 - Conveyor 22 - Transfering

      A     "M 87.1";
      AN    "M 87.2";
      A     "M 82.0";
      A     "M 83.2";
      S     "M 83.3";
NETWORK
TITLE =Step 23N5 - Conveyor 22 - Steps Register - Reset

      A(    ;
      O     "B 15.7";
      O     "Timer 83";
      )     ;
      A     "M 82.0";
      A     "M 83.3";
      S     "M 83.4";
NETWORK
TITLE =Conveyor  22 VFD - Release

      A(    ;
      A     "M 83.1";
      AN    "M 83.2";
      O     ;
      A     "M 83.3";
      AN    "M 83.4";
      )     ;
      A     "M 82.0";
      AN    "M 11.1"; // VFD NOT All Ready !
      =     "A 53.6";
      =     "A 53.7";
END_FUNCTION

FUNCTION "CONVEYOR 23 - DELIV. HI" : VOID
TITLE =Conveyor 23 - Delivery Second Level
//
NAME : POS_15_H
VERSION : 0.0


VAR_TEMP
  MAIN_SERVICE_2_SW : BOOL ;
  SERVICE_RUN : BOOL ;
END_VAR
BEGIN
NETWORK
TITLE =Conveyor 23 - Service

      A     "HMI_DB".ALL_SERVICE_ENABLE_SW;
      A     "HMI_DB".CONVEYOR_21_SERVICE_SW;
      A     "HMI_DB".SERVICE_SW_2_STATUS;
      =     #MAIN_SERVICE_2_SW;
//;
      A     #MAIN_SERVICE_2_SW;
      O     "M 86.1";
      JNB   CO23;
//;
      A     "HMI_DB".HMI_CONVEYOR_23_TEST_SSW;
      =     #SERVICE_RUN;
//;
      AN    #MAIN_SERVICE_2_SW;
      R     "HMI_DB".HMI_CONVEYOR_23_TEST_SSW;

CO23: R     #SERVICE_RUN;
      FP    "FP 149.3";
      =     "M 86.1";
NETWORK
TITLE =Delivery Conveyor 23 - Running TimeOut  30s
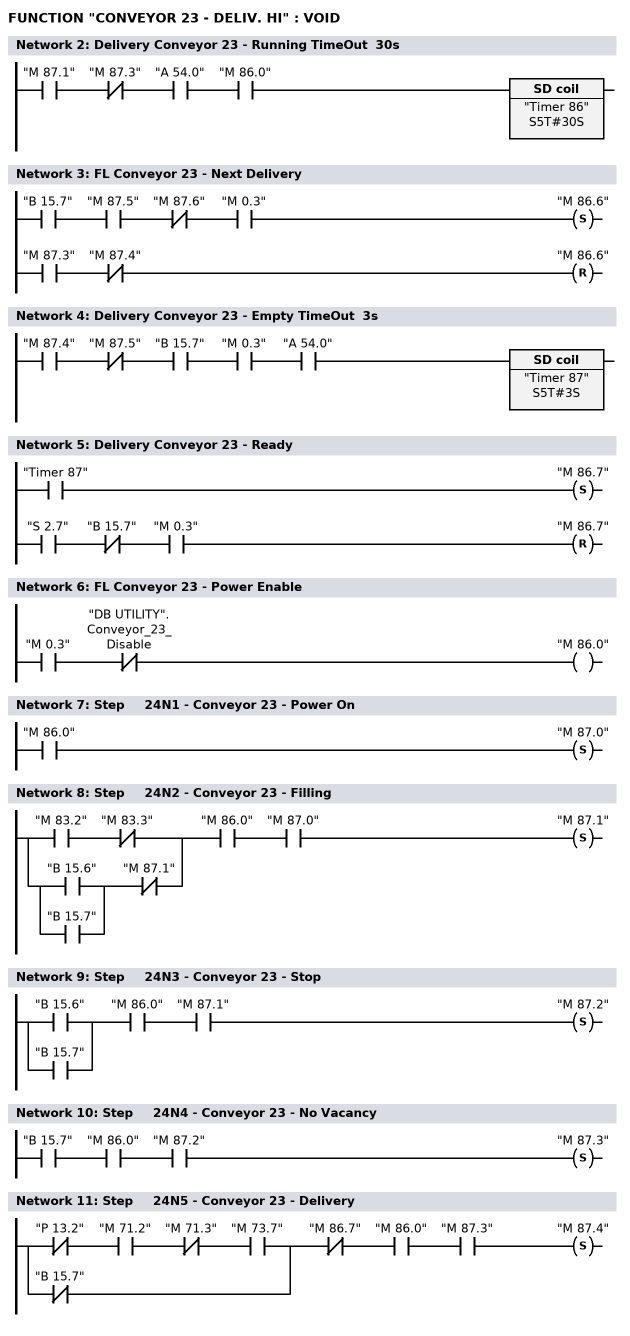

      A     "M 87.1";
      AN    "M 87.3";
      A     "A 54.0";
      A     "M 86.0";
      L     S5T#30S;
      SD    "Timer 86";
NETWORK
TITLE =FL Conveyor 23 - Next Delivery

      A     "B 15.7";
      A     "M 87.5";
      AN    "M 87.6";
      A     "M 0.3";
      S     "M 86.6";
//;
      A     "M 87.3";
      AN    "M 87.4";
      R     "M 86.6";
NETWORK
TITLE =Delivery Conveyor 23 - Empty TimeOut  3s

      A     "M 87.4";
      AN    "M 87.5";
      A     "B 15.7";
      A     "M 0.3";
      A     "A 54.0";
      L     S5T#3S;
      SD    "Timer 87";
NETWORK
TITLE =Delivery Conveyor 23 - Ready

      A     "Timer 87";
      S     "M 86.7";
//;
      A     "S 2.7";
      AN    "B 15.7";
      A     "M 0.3";
      R     "M 86.7";
NETWORK
TITLE =FL Conveyor 23 - Power Enable

      A     "M 0.3";
      AN    "DB UTILITY".Conveyor_23_Disable;
      =     "M 86.0";
NETWORK
TITLE =Step     24N1 - Conveyor 23 - Power On

      A     "M 86.0";
      S     "M 87.0";
NETWORK
TITLE =Step     24N2 - Conveyor 23 - Filling

      A(    ;
      A     "M 83.2";
      AN    "M 83.3";
      O     ;
      A(    ;
      O     "B 15.6";
      O     "B 15.7";
      )     ;
//      O     #SERVICE_RUN
      AN    "M 87.1";
      )     ;
      A     "M 86.0";
      A     "M 87.0";
      S     "M 87.1";
NETWORK
TITLE =Step     24N3 - Conveyor 23 - Stop

      A(    ;
      O     "B 15.6";
      O     "B 15.7";
      )     ;
      A     "M 86.0";
      A     "M 87.1";
      S     "M 87.2";
NETWORK
TITLE =Step     24N4 - Conveyor 23 - No Vacancy

      A     "B 15.7";
      A     "M 86.0";
      A     "M 87.2";
      S     "M 87.3";
NETWORK
TITLE =Step     24N5 - Conveyor 23 - Delivery

      A(    ;
      AN    "P 13.2";
      A     "M 71.2";
      AN    "M 71.3";
      A     "M 73.7";
      ON    "B 15.7";
      )     ;
      AN    "M 86.7";
      A     "M 86.0";
      A     "M 87.3";
      S     "M 87.4";
NETWORK
TITLE =Write 1 to Steps 0-3 Byte Register MB87

      A(    ;
      O     "M 86.6";
      O     "M 86.7";
      )     ;
      A     "M 87.4";
      A     "M 86.0";
      JC    M001;
      JU    M002;

M001: L     2#1111;
      T     "MB 87";

M002: NOP   0;
NETWORK
TITLE =Step     24N6 - Conveyor 23 - Delivery Done
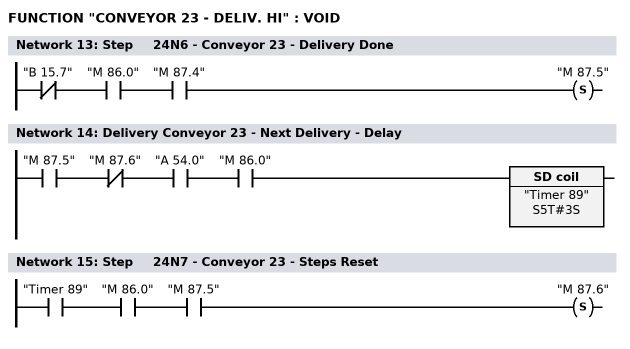

      AN    "B 15.7";
      A     "M 86.0";
      A     "M 87.4";
      S     "M 87.5";
NETWORK
TITLE =Delivery Conveyor 23 - Next Delivery - Delay

      A     "M 87.5";
      AN    "M 87.6";
      A     "A 54.0";
      A     "M 86.0";
      L     S5T#3S;
      SD    "Timer 89";
NETWORK
TITLE =Step     24N7 - Conveyor 23 - Steps Reset

      A     "Timer 89";
      A     "M 86.0";
      A     "M 87.5";
      S     "M 87.6";
NETWORK
TITLE =Steps Register - Reset

      A(    ;
      O     "M 87.6";
      O     "Timer 86";
      )     ;
      A     "M 86.0";
      JC    M003;
      JU    M004;

M003: L     2#0;
      T     "MW 87";

M004: NOP   0;
NETWORK
TITLE =Conveyor  23 VFD - Release
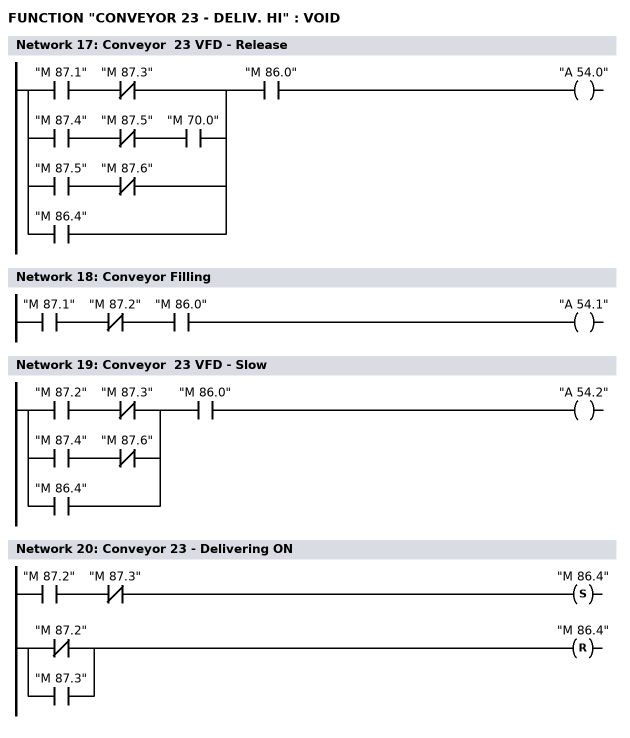

      A(    ;
      A     "M 87.1";
      AN    "M 87.3";
      O     ;
      A     "M 87.4";
      AN    "M 87.5";
      A     "M 70.0";
      O     ;
      A     "M 87.5";
      AN    "M 87.6";
      O     "M 86.4";
      )     ;
      A     "M 86.0";
      =     "A 54.0";
NETWORK
TITLE =Conveyor Filling

      A     "M 87.1";
      AN    "M 87.2";
      A     "M 86.0";
      =     "A 54.1";
NETWORK
TITLE =Conveyor  23 VFD - Slow

      A(    ;
      A     "M 87.2";
      AN    "M 87.3";
      O     ;
      A     "M 87.4";
      AN    "M 87.6";
      O     "M 86.4";
      )     ;
      A     "M 86.0";
      =     "A 54.2";
NETWORK
TITLE =Conveyor 23 - Delivering ON

      A     "M 87.2";
      AN    "M 87.3";
      S     "M 86.4";
      A(    ;
      ON    "M 87.2";
      O     "M 87.3";
      )     ;
      R     "M 86.4";
END_FUNCTION

FUNCTION "LIGHT BAR" : VOID
TITLE =Light Bar
VERSION : 0.1


VAR_TEMP
  BARRIER_BLINKER : BOOL ;	//Feeder Safety Light Barrier
  STATUS_BLANKER : BOOL ;
  CLEARING_BLINKER : BOOL ;
END_VAR
BEGIN
NETWORK
TITLE =Light Barrier - Blinker
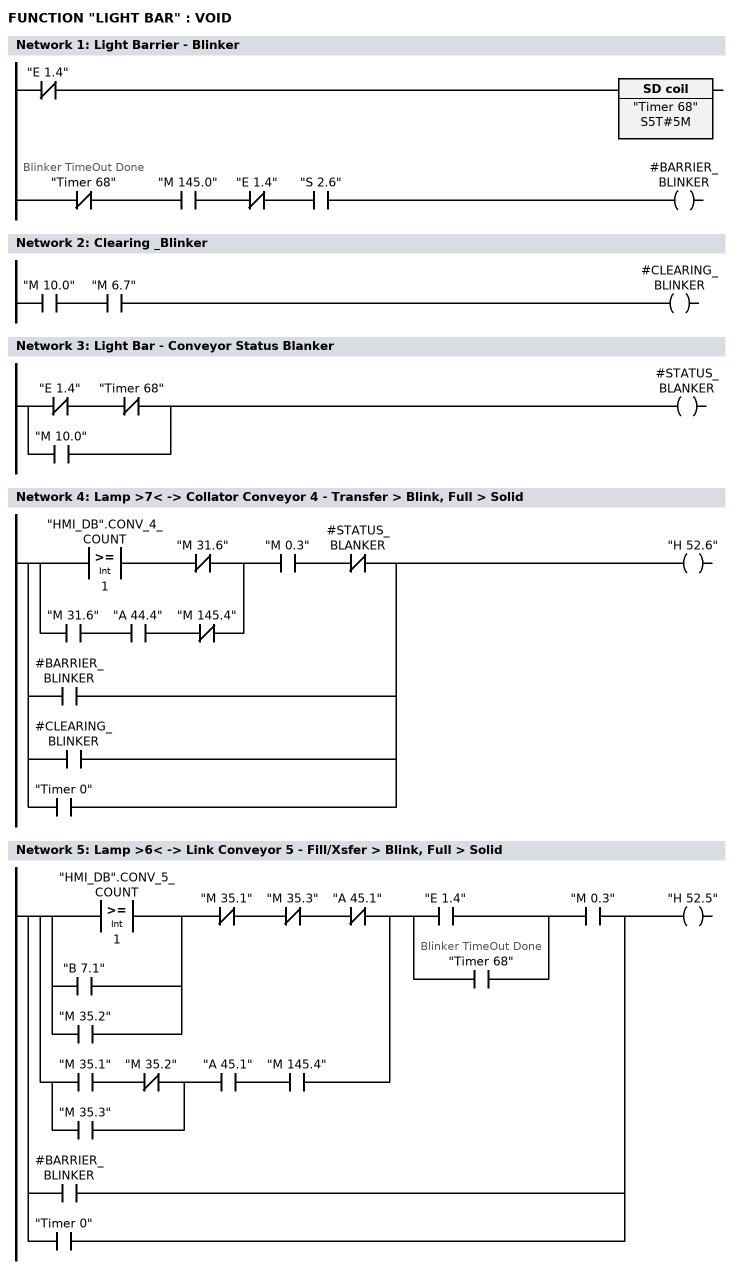

      ON    "E 1.4";
      L     S5T#5M;
      SD    "Timer 68"; // Blinker TimeOut Start
//;
      A(    ;
      AN    "Timer 68"; // Blinker TimeOut Done
      A     "M 145.0";
      )     ;
      AN    "E 1.4";
      A     "S 2.6";
      =     #BARRIER_BLINKER;
NETWORK
TITLE =Clearing _Blinker

      A     "M 10.0";
      A     "M 6.7";
      =     #CLEARING_BLINKER;
NETWORK
TITLE =Light Bar - Conveyor Status Blanker

      AN    "E 1.4";
      AN    "Timer 68";
      O     "M 10.0";
      =     #STATUS_BLANKER;
NETWORK
TITLE =Lamp >7< -> Collator Conveyor 4 - Transfer > Blink, Full > Solid

      A(    ;

      A(    ; // Solid
      A(    ;
      L     "HMI_DB".CONV_4_COUNT;
      L     1;
      >=I   ;
      )     ;
      AN    "M 31.6";
      )     ; // Solid

      O     ;

      A(    ; // Blink
      A     "M 31.6";
      A     "A 44.4";
      AN    "M 145.4";
      )     ; // Blink

      )     ;
      A     "M 0.3";
      AN    #STATUS_BLANKER;
      O     #BARRIER_BLINKER;
      O     #CLEARING_BLINKER;
      O     "Timer 0";
      =     "H 52.6";
NETWORK
TITLE =Lamp >6< -> Link Conveyor 5 - Fill/Xsfer > Blink, Full > Solid

      A(    ;

      A(    ; // Solid
      A(    ;
      A(    ;
      L     "HMI_DB".CONV_5_COUNT;
      L     1;
      >=I   ;
      )     ;
      O     "B 7.1";
      )     ;
      O     "M 35.2";
      AN    "M 35.1";
      AN    "M 35.3";
      AN    "A 45.1";
      )     ; // Solid

      O     ;

      A(    ; // Blink
      A(    ;
      A     "M 35.1";
      AN    "M 35.2";
      O     ;
      A     "M 35.3";
      )     ;
      A     "A 45.1";
      A     "M 145.4";
      )     ; // Blink

      )     ;
      A(    ;
      A     "E 1.4";
      O     "Timer 68"; // Blinker TimeOut Done
      )     ;
      A     "M 0.3";
      O     #BARRIER_BLINKER;
      O     "Timer 0";
      =     "H 52.5";
NETWORK
TITLE =Lamp >5< -> Delivery Conveyor 6 - Fill > Blink, Full > Solid

      A(    ;

      A(    ; // Solid
      A(    ;
      A(    ;
      L     "HMI_DB".CONV_6_COUNT;
      L     1;
      >=I   ;
      )     ;
      O     "B 7.2";
      )     ;
      O     "M 39.2";
      AN(   ;
      A     "M 39.1";
      AN    "M 39.2";
      )     ;
      AN    "A 45.4";
      )     ; // Solid

      O     ;

      A(    ; // Blink
      A     "M 39.1";
      AN    "M 39.2";
      A     "A 45.4";
      AN    "M 145.4";
      )     ; // Blink

      )     ;
      A(    ;
      A     "E 1.4";
      O     "Timer 68"; // Blinker TimeOut Done
      )     ;
      A     "M 0.3";
      O     #BARRIER_BLINKER;
      O     "Timer 0";
      =     "H 52.4";
NETWORK
TITLE =Lamp >4< -> Pivot 10 -> 11L/21H - Fill > Blink, Full > Solid
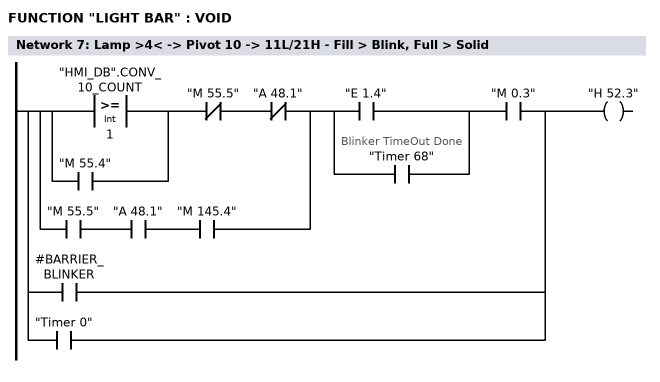

      A(    ;

      A(    ; // Solid
      A(    ;
      L     "HMI_DB".CONV_10_COUNT;
      L     1;
      >=I   ;
      )     ;
      O     "M 55.4";
      AN    "M 55.5";
      AN    "A 48.1";
      )     ; // Solid

      O     ;

      A(    ; // Blink
      A     "M 55.5";
      A     "A 48.1";
      A     "M 145.4";
      )     ; // Blink

      )     ;
      A(    ;
      A     "E 1.4";
      O     "Timer 68"; // Blinker TimeOut Done
      )     ;
      A     "M 0.3";
      O     #BARRIER_BLINKER;
      O     "Timer 0";
      =     "H 52.3";
NETWORK
TITLE =Lamp >3< -> Link Conveyors 11L/21H - Fill > Blink, Full > Solid

      A(    ;

      A(    ; // Solid
      A(    ;
      A(    ;
      A(    ;
      L     "HMI_DB".CONV_11_COUNT;
      L     "HMI_DB".CONV_21_COUNT;
      +I    ;
      L     1;
      >=I   ;
      )     ;
      O     "B 10.7";
      O     "B 15.4";
      )     ;
      O     "M 59.2";
      O     "M 79.2";
      )     ;
      AN(   ;
      A     "M 59.1";
      AN    "M 59.2";
      )     ;
      AN(   ;
      A     "M 79.1";
      AN    "M 79.2";
      )     ;
      AN    "M 59.3";
      AN    "M 79.3";
      AN    "A 48.3";
      AN    "A 53.4";
      )     ; // Solid

      O     ;

      A(    ; // Blink
      A(    ;
      A(    ;
      A     "M 59.1";
      AN    "M 59.2";
      O     ;
      A     "M 79.1";
      AN    "M 79.2";
      )     ;
      O     ;
      A(    ;
      A     "M 59.3";
      O     "M 79.3";
      )     ;
      )     ;
      A(    ;
      O     "A 48.3";
      O     "A 53.4";
      )     ;
      AN    "M 145.4";
      )     ; // Blink

      )     ;
      A(    ;
      A     "E 1.4";
      O     "Timer 68"; // Blinker TimeOut Done
      )     ;
      A     "M 0.3";
      O     #BARRIER_BLINKER;
      O     "Timer 0";
      =     "H 52.2";

NETWORK
TITLE =Lamp >2< -> Link Conveyors 12L/22H - Fill > Blink, Full > Solid

      A(    ;

      A(    ; // Solid
      A(    ;
      A(    ;
      A(    ;
      L     "HMI_DB".CONV_12_COUNT;
      L     "HMI_DB".CONV_22_COUNT;
      +I    ;
      L     1;
      >=I   ;
      )     ;
      O     "B 11.0";
      O     "B 15.5";
      )     ;
      O     "M 63.2";
      O     "M 83.2";
      )     ;
      AN(   ;
      A     "M 63.1";
      AN    "M 63.2";
      )     ;
      AN(   ;
      A     "M 83.1";
      AN    "M 83.2";
      )     ;
      AN    "M 63.3";
      AN    "M 83.3";
      AN    "A 48.6";
      AN    "A 53.6";
      )     ; // Solid

      O     ;

      A(    ; // Blink
      A(    ;
      A(    ;
      A     "M 63.1";
      AN    "M 63.2";
      O     ;
      A     "M 83.1";
      AN    "M 83.2";
      )     ;
      O     ;
      A(    ;
      A     "M 63.3";
      O     "M 83.3";
      )     ;
      )     ;
      A(    ;
      O     "A 48.6";
      O     "A 53.6";
      )     ;
      A     "M 145.4";
      )     ; // Blink

      )     ;
      A(    ;
      A     "E 1.4";
      O     "Timer 68"; // Blinker TimeOut Done
      )     ;
      A     "M 0.3";
      O     #BARRIER_BLINKER;
      O     "Timer 0";
      =     "H 52.1";

NETWORK
TITLE =Lamp >1< -> Output Conveyors 13L/23H - Fill > Blink,Full > Solid

      A(    ; // Solid

      A(    ;
      L     "HMI_DB".CONV_13_COUNT;
      L     "HMI_DB".CONV_23_COUNT;
      +I    ;
      L     1;
      >=I   ;
      )     ;
      O     "B 11.2";
      O     "B 15.7";
      )     ; // Solid

      A(    ;
      A     "E 1.4";
      O     "Timer 68"; // Blinker TimeOut Done
      )     ;
      A     "M 0.3";
      AN    #STATUS_BLANKER;
      O     #BARRIER_BLINKER;
      O     #CLEARING_BLINKER;
      O     "Timer 0";
      =     "H 52.0";
END_FUNCTION

FUNCTION "HMI CONTROL" : VOID
TITLE =HMI Control - Screen 0 SSW Inputs
//Screen 0 - "RUN" Screen
NAME : HMI_CTRL
VERSION : 0.1


VAR_TEMP
  SERVICE_ON : BOOL ;
  CLEARING_ON : BOOL ;
  HAND_FEED : BOOL ;
  UPDATE_PULSE : BOOL ;
END_VAR
BEGIN
NETWORK
TITLE =New HMI Panel Switches
